DATA_BLOCK "Sim"
TITLE = 'Instance of the plant simulation'
{ S7_Optimized_Access := 'TRUE' }
VERSION : 0.1
NON_RETAIN
"FB_ProcessSim"

BEGIN

END_DATA_BLOCK
